Universal Robots URScript: EdgeProg.script

def EdgeProg():
  # Global parameters:
  global speed_ms    = 0.250
  global speed_rads  = 0.750
  global accel_mss   = 1.200
  global accel_radss = 1.200
  global blend_radius_m = 0.001
  global ref_frame = p[0,0,0,0,0,0]

  #
  # TO REMOVE HEADER:
  # Go to "Program" -> "Post-Processor Editor"
  # Select "Universal Robots"
  # Set "INCLUDE_HEADER" to "False"
  #
  #--------------------------
  # Add any default subprograms here
  # For example, to drive a gripper as a program call:
  # def Gripper_Open():
  #   ...
  # end
  #
  # Example to drive a spray gun:
  def SprayOn(value):
    # use the value as an output:
    DO_SPRAY = 5
    if value == 0:
      set_standard_digital_out(DO_SPRAY, False)
    else:
      set_standard_digital_out(DO_SPRAY, True)
    end
  end

  # Example to drive an extruder:
  def Extruder(value):
    # use the value as an output:
    if value < 0:
      # stop extruder
    else:
      # start extruder
    end
  end

  # Example to move an external axis
  def MoveAxis(value):
    # use the value as an output:
    DO_AXIS_1 = 1
    DI_AXIS_1 = 1
    if value <= 0:
      set_standard_digital_out(DO_AXIS_1, False)

      # Wait for digital input to change state
      #while (get_standard_digital_in(DI_AXIS_1) != False):
      #  sync()
      #end
    else:
      set_standard_digital_out(DO_AXIS_1, True)

      # Wait for digital input to change state
      #while (get_standard_digital_in(DI_AXIS_1) != True):
      #  sync()
      #end
    end
  end
  #--------------------------


  # Main program:
  # Program generated by RoboDK v6.0.7 for UR10 on XX/XX/XXXX 18:00:00
  # Using nominal kinematics.
  ref_frame = p[0.100500, -0.200250, 0.300125, 0.547381, -0.295318, 0.260260]
  set_tcp(p[-0.001500, 0.002250, 0.099875, -1.759988, 1.759988, 0.729011])
  speed_ms    = 0.123
  speed_rads  = 0.582
  blend_radius_m = 0.000
  movej([-0.087266, -0.087266, 0.261799, 0.174533, 0.698132, -0.174533],accel_radss,speed_rads,t=0,r=0)
  blend_radius_m = 0.013
  movel(pose_trans(ref_frame,p[-0.624230, 0.571208, 0.454620, -0.100914, 1.591504, -1.158572]),accel_mss,speed_ms,t=0,r=0.013)
  halt() # reimplement this function to force stop
  sleep(1.234)
  popup("A long message with "quotes", 'apostrophes' & symbols: <>[]{}()=+-*/%;#@! and more text to make it longer than eighty characters","Message",False,False,blocking=True)
  # Comment with ; semicolon
  Gripper = ON
  set_tool_digital_out(2, False)
  Pressure = 0.75
  while (PartPresent != True):
    sync()
  end
  while (get_standard_digital_in(7) != 1):
    sync()
  end
  DoSomething(1, 2)
  x = 1
  movej([0.349066, -0.174533, 0.349066, 0.000000, 0.523599, 0.000000],accel_radss,speed_rads,t=0,r=0)
  # End of main program
end

EdgeProg()
